TYPE "DT_MEASUREMENT_ALL"
VERSION : 0.1
   STRUCT
      TURBINE_AND_HPU : "DT_MEASUREMENT_SYSTEM_TURBINE_AND_HPU";
      GENERATOR_MECHANICAL : "DT_MEASUREMENT_SYSTEM_GENERATOR_MECHANICAL";
      GENERATOR_MEASUREMENT : "DT_MEASUREMENT_SYSTEM_GENERATOR_MEASUREMENT";
      GENERATOR_PROTECTION : "DT_MEASUREMENT_SYSTEM_GENERATOR_PROTECTION";
      GENERATOR_EXCITATION : "DT_MEASUREMENT_SYSTEM_GENERATOR_EXCITATION";
      LINE_MEAS_DEVICE : "DT_MEASUREMENT_SYSTEM_LINE_MEAS";
      TRAFO_PROTECTION : "DT_MEASUREMENT_SYSTEM_LINE_PROTECTION";
      CONTROL : "DT_MEASUREMENT_SYSTEM_CONTROL";
      CWS_AND_LOU : "DT_MEASUREMENT_SYSTEM_CWS_AND_LOU";
      AUX_SUPPLY : "DT_MEASUREMENT_SYSTEM_AUX_SUPPLY";
      TRAFO_AND_OTHER : "DT_MEASUREMENT_SYSTEM_TRAFO_AND_OTHER";
      SPARE : "DT_MEASUREMENT_SYSTEM_SPARE";
   END_STRUCT;

END_TYPE

